INTERFACE I_OtlpValue

PROPERTY eType : E_ValueType
GET
END_GET
END_PROPERTY

// deallocates all data owned by the value without deleting the object itself.
METHOD free
END_METHOD

END_INTERFACE

(* stored: Version 1.1.0.1
   Itf I_OtlpValue: Id {fc55bdb3-176f-48d0-b16b-8f81387d6392}
   Property eType: Id {f215879f-eadf-4cab-a2f7-31f77a67d6d2}
   Get Get: Id {bdc18bae-f138-4217-a020-1f99bbb64531}
   Method free: Id {063e0f66-c6cb-45a4-a9ca-6cfd5e61a0ea} *)
